FUNCTION_BLOCK F (* Needs reading R1: a variable stepped by +1 and dispatched from two control states. It may be a step number or a count *)
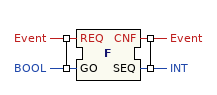
  EVENT_INPUT
    REQ WITH GO;
  END_EVENT
  EVENT_OUTPUT
    CNF WITH SEQ;
  END_EVENT
  VAR_INPUT
    GO : BOOL;
  END_VAR
  VAR_OUTPUT
    SEQ : INT;
  END_VAR
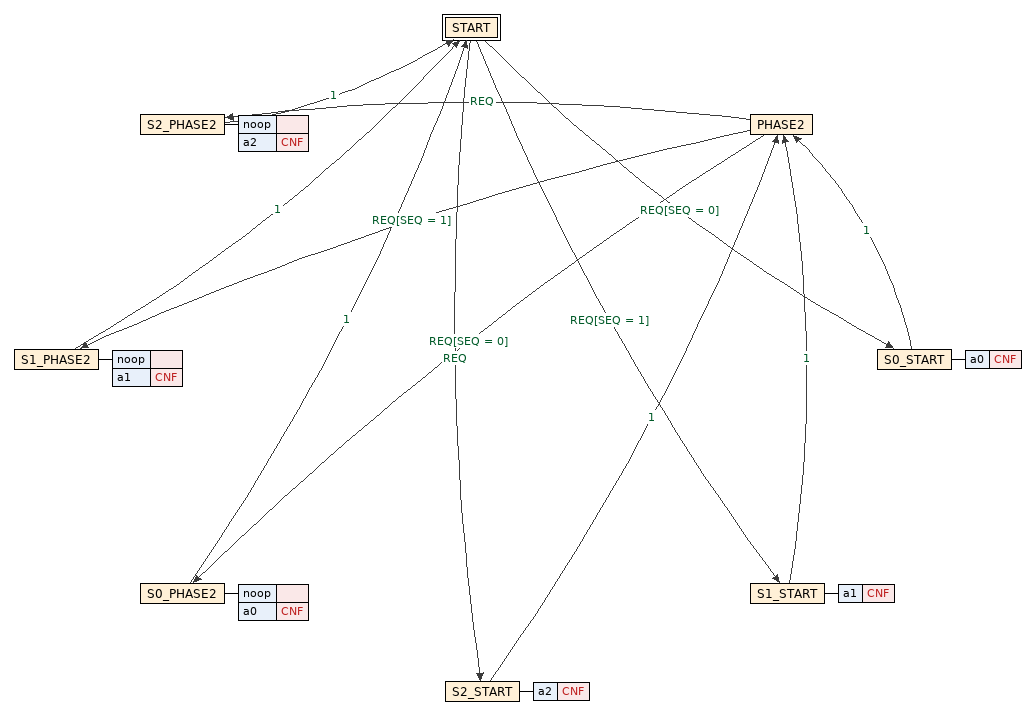
  EC_STATES
    START;
    PHASE2;
    S0_START : a0 -> CNF;
    S1_START : a1 -> CNF;
    S2_START : a2 -> CNF;
    S0_PHASE2 : noop, a0 -> CNF;
    S1_PHASE2 : noop, a1 -> CNF;
    S2_PHASE2 : noop, a2 -> CNF;
  END_STATES
  EC_TRANSITIONS
    START TO S0_START := REQ[SEQ = 0];
    START TO S1_START := REQ[SEQ = 1];
    START TO S2_START := REQ;
    PHASE2 TO S0_PHASE2 := REQ[SEQ = 0];
    PHASE2 TO S1_PHASE2 := REQ[SEQ = 1];
    PHASE2 TO S2_PHASE2 := REQ;
    S0_START TO PHASE2 := 1;
    S1_START TO PHASE2 := 1;
    S2_START TO PHASE2 := 1;
    S0_PHASE2 TO START := 1;
    S1_PHASE2 TO START := 1;
    S2_PHASE2 TO START := 1;
  END_TRANSITIONS
  ALGORITHM a0 IN ST:
IF GO THEN
  SEQ := SEQ + 1;
END_IF;
  END_ALGORITHM
  ALGORITHM a1 IN ST:
SEQ := SEQ + 1;
  END_ALGORITHM
  ALGORITHM a2 IN ST:
SEQ := 0;
  END_ALGORITHM
  ALGORITHM noop IN ST:
SEQ := SEQ;
  END_ALGORITHM
END_FUNCTION_BLOCK
